SYSTEM Adaptive_Identification (* Offline only; native export and runtime validation pending *)
  APPLICATION Identification_Offline
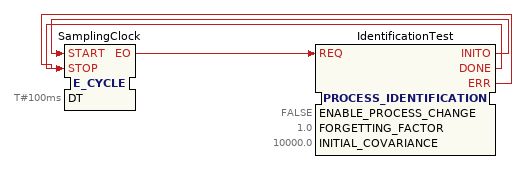
    FBS
      SamplingClock : E_CYCLE(DT := T#100ms);
      IdentificationTest : PROCESS_IDENTIFICATION(ENABLE_PROCESS_CHANGE := FALSE, FORGETTING_FACTOR := 1.0, INITIAL_COVARIANCE := 10000.0);
    END_FBS
    EVENT_CONNECTIONS
      IdentificationTest.INITO TO SamplingClock.START;
      SamplingClock.EO TO IdentificationTest.REQ;
      IdentificationTest.DONE TO SamplingClock.STOP;
      IdentificationTest.ERR TO SamplingClock.STOP;
    END_CONNECTIONS
  END_APPLICATION
  DEVICE LocalIdentification : FORTE_PC(MGR_ID := "localhost:61499")
    {SET_ATTRIBUTE(Profile, HOLOBLOC)} (* device profile *)
    RESOURCE EMB_RES : EMB_RES
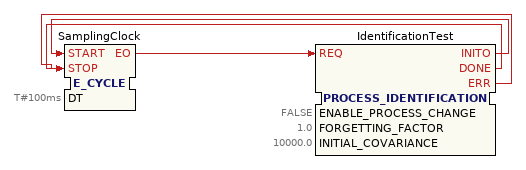
      FBS
        IdentificationTest : PROCESS_IDENTIFICATION(ENABLE_PROCESS_CHANGE := FALSE, FORGETTING_FACTOR := 1.0, INITIAL_COVARIANCE := 10000.0);
        SamplingClock : E_CYCLE(DT := T#100ms);
      END_FBS
      EVENT_CONNECTIONS
        IdentificationTest.INITO TO SamplingClock.START;
        IdentificationTest.DONE TO SamplingClock.STOP;
        IdentificationTest.ERR TO SamplingClock.STOP;
        SamplingClock.EO TO IdentificationTest.REQ;
      END_CONNECTIONS
    END_RESOURCE
  END_DEVICE
  MAPPINGS
    Identification_Offline.IdentificationTest ON LocalIdentification.EMB_RES.IdentificationTest;
    Identification_Offline.SamplingClock ON LocalIdentification.EMB_RES.SamplingClock;
  END_MAPPINGS
END_SYSTEM
